(* IEC 61131-3 sources: Simulierte-Foerderanlagensteuerung/plc/function_blocks, 6 files *)

(* ---- FB_Alarm.st ---- *)
(* ============================================================================
   FB_Alarm.st
   Störmeldespeicher, Priorisierung und First-out-Erkennung.

   - Ueberlast und Not-Halt sind "lebende" Bedingungen (fallen mit dem Signal).
   - Timeout-/Stau-/Sensorstoerungen werden gespeichert und nur quittiert,
     wenn die Ursache nicht mehr ansteht.
   - eFirst haelt die zuerst aufgetretene Stoerung fest.
   ============================================================================ *)

FUNCTION_BLOCK FB_Alarm
VAR_INPUT
    xOverload            : BOOL;
    xEmergency           : BOOL;
    xStartTimeout        : BOOL;
    xStopTimeout         : BOOL;
    xJam                 : BOOL;
    xSensorInconsistency : BOOL;
    xReset               : BOOL;
END_VAR
VAR_OUTPUT
    eActive    : E_FaultCode;
    eFirst     : E_FaultCode;
    xAnyFault  : BOOL;
    xLampRed   : BOOL;
    xLampYellow: BOOL;
    xBuzzer    : BOOL;
    xOverloadLatched  : BOOL;
    xEmergencyLatched : BOOL;
    xStartLatched     : BOOL;
    xStopLatched      : BOOL;
    xJamLatched       : BOOL;
    xSensorLatched    : BOOL;
END_VAR

    (* --- Ereignisstoerungen speichern --- *)
    IF xOverload THEN
        xOverloadLatched := TRUE;
    END_IF;
    IF xEmergency THEN
        xEmergencyLatched := TRUE;
    END_IF;
    IF xStartTimeout THEN
        xStartLatched := TRUE;
    END_IF;
    IF xStopTimeout THEN
        xStopLatched := TRUE;
    END_IF;
    IF xJam THEN
        xJamLatched := TRUE;
    END_IF;
    IF xSensorInconsistency THEN
        xSensorLatched := TRUE;
    END_IF;

    (* --- Sammelstoerung --- *)
    xAnyFault := xOverloadLatched
                 OR xEmergencyLatched
                 OR xStartLatched
                 OR xStopLatched
                 OR xJamLatched
                 OR xSensorLatched;

    (* --- Quittung nur, wenn keine Ursache mehr ansteht --- *)
    IF xReset
       AND NOT xOverload
       AND NOT xEmergency
       AND NOT xStartTimeout
       AND NOT xStopTimeout
       AND NOT xJam
       AND NOT xSensorInconsistency THEN
        xOverloadLatched := FALSE;
        xEmergencyLatched := FALSE;
        xStartLatched := FALSE;
        xStopLatched := FALSE;
        xJamLatched := FALSE;
        xSensorLatched := FALSE;
    END_IF;

    (* --- Priorisierte Anzeige der aktiven Stoerung --- *)
    IF xEmergencyLatched THEN
        eActive := E_FaultCode.FAULT_EMERGENCY;
    ELSIF xOverloadLatched THEN
        eActive := E_FaultCode.FAULT_OVERLOAD;
    ELSIF xStartLatched THEN
        eActive := E_FaultCode.FAULT_START_TIMEOUT;
    ELSIF xStopLatched THEN
        eActive := E_FaultCode.FAULT_STOP_TIMEOUT;
    ELSIF xJamLatched THEN
        eActive := E_FaultCode.FAULT_JAM;
    ELSIF xSensorLatched THEN
        eActive := E_FaultCode.FAULT_SENSOR_INCONSISTENCY;
    ELSE
        eActive := E_FaultCode.FAULT_NONE;
    END_IF;

    (* --- First-out --- *)
    IF (eFirst = E_FaultCode.FAULT_NONE) AND xAnyFault THEN
        eFirst := eActive;
    END_IF;
    IF xReset AND NOT xAnyFault THEN
        eFirst := E_FaultCode.FAULT_NONE;
    END_IF;

    (* --- Meldeorgane --- *)
    xLampRed := xAnyFault;
    xBuzzer := xAnyFault;
    xLampYellow := (eActive = E_FaultCode.FAULT_JAM)
                   OR (eActive = E_FaultCode.FAULT_SENSOR_INCONSISTENCY);
END_FUNCTION_BLOCK

(* ---- FB_ConveyorProcess.st ---- *)
(* ============================================================================
   FB_ConveyorProcess.st
   Prozessablauf Automatikbetrieb.

   Zwei Varianten, gesteuert durch die Konstante AUTO_CONTINUOUS:
     - Bedarfsbetrieb (FALSE): Start bei Werkstueck am Einlauf, Nachlauf nach
       dem Auslauf, dann Rueckkehr nach IDLE.
     - Dauerlauf (TRUE): Start beim Aktivieren der Automatik, kein Stopp.

   Ausgaenge sind Impulse (ein Zyklus) fuer die Motorsteuerung.
   ============================================================================ *)

FUNCTION_BLOCK FB_ConveyorProcess
VAR_INPUT
    xEnable      : BOOL;   (* Automatik aktiv, READY, keine Stoerung *)
    xEntrySensor : BOOL;   (* B1 *)
    xExitSensor  : BOOL;   (* B2 *)
END_VAR
VAR_OUTPUT
    xStartPulse : BOOL;    (* Startimpuls an Motorsteuerung *)
    xStopPulse  : BOOL;    (* Stopimpuls an Motorsteuerung *)
    eState      : E_ProcessState;
END_VAR
VAR
    xEnablePrev : BOOL;
    tonRunOn    : TON;
    xRunOnCond  : BOOL;
END_VAR

    xStartPulse := FALSE;
    xStopPulse  := FALSE;

    (* Nachlauf-Timer jede Scan aufrufen; ausserhalb P_RUN_ON zuruecksetzen *)
    xRunOnCond := (eState = E_ProcessState.P_RUN_ON) AND NOT xExitSensor;
    tonRunOn(IN := xRunOnCond, PT := T_RUN_ON);

    IF NOT xEnable THEN
        IF xEnablePrev THEN
            xStopPulse := TRUE;   (* Automatik verlassen -> Band stoppen *)
        END_IF;
        eState := E_ProcessState.P_IDLE;
        xEnablePrev := FALSE;
    ELSE
        CASE eState OF
            E_ProcessState.P_IDLE :
                IF AUTO_CONTINUOUS THEN
                    IF NOT xEnablePrev THEN
                        xStartPulse := TRUE;
                    END_IF;
                    eState := E_ProcessState.P_TRANSPORT;
                ELSE
                    IF xEntrySensor THEN
                        xStartPulse := TRUE;
                        eState := E_ProcessState.P_TRANSPORT;
                    END_IF;
                END_IF;

            E_ProcessState.P_TRANSPORT :
                IF (NOT AUTO_CONTINUOUS) AND xExitSensor THEN
                    eState := E_ProcessState.P_RUN_ON;
                END_IF;

            E_ProcessState.P_RUN_ON :
                IF tonRunOn.Q THEN
                    xStopPulse := TRUE;
                    eState := E_ProcessState.P_IDLE;
                END_IF;

            ELSE
                eState := E_ProcessState.P_IDLE;
        END_CASE;
        xEnablePrev := TRUE;
    END_IF;
END_FUNCTION_BLOCK

(* ---- FB_Counter.st ---- *)
(* ============================================================================
   FB_Counter.st
   Werkstueckzaehlung.

   Gezaehlt wird am Auslauf ueber die steigende Flanke des Sensors B2.
   Begruendung: Der Auslauf repraesentiert ein fertig transportiertes Werkstueck.
   Die Flankenauswertung (R_TRIG) verhindert Mehrfachzaehlung, solange der
   Sensor aktiv bleibt.
   ============================================================================ *)

FUNCTION_BLOCK FB_Counter
VAR_INPUT
    xExitSensor : BOOL;    (* B2 *)
    xResetCount : BOOL;
END_VAR
VAR_OUTPUT
    diCount      : DINT;
    xJustCounted : BOOL;   (* Impuls fuer HMI/Statistik *)
END_VAR
VAR
    rtrigExit : R_TRIG;
END_VAR

    rtrigExit(CLK := xExitSensor);
    xJustCounted := FALSE;

    IF rtrigExit.Q THEN
        diCount := diCount + 1;
        xJustCounted := TRUE;
    END_IF;

    IF xResetCount THEN
        diCount := 0;
    END_IF;
END_FUNCTION_BLOCK

(* ---- FB_JamDetection.st ---- *)
(* ============================================================================
   FB_JamDetection.st
   Stau-/Blockadeerkennung.

   Verfahren: Ein Werkstueck wird am Einlauf erkannt und der Antrieb laeuft.
   Erreicht es den Auslauf nicht innerhalb T_MAX_TRANSPORT, liegt ein Stau vor.
   Die Stau-Stoerung wird bis zur Quittung gespeichert.
   ============================================================================ *)

FUNCTION_BLOCK FB_JamDetection
VAR_INPUT
    xEntrySensor      : BOOL;   (* B1 *)
    xExitSensor       : BOOL;   (* B2 *)
    xConveyorRun      : BOOL;   (* Antrieb angesteuert bzw. laeuft *)
    xReset            : BOOL;
END_VAR
VAR_OUTPUT
    xJam              : BOOL;
    xTransportPending : BOOL;   (* Werkstueck unterwegs, Auslauf erwartet *)
END_VAR
VAR
    rtrigEntry : R_TRIG;
    tonJam     : TON;
END_VAR

    rtrigEntry(CLK := xEntrySensor);

    (* Transportauftrag setzen, sobald ein Werkstueck einlaeuft und der Antrieb laeuft *)
    IF rtrigEntry.Q AND xConveyorRun THEN
        xTransportPending := TRUE;
    END_IF;

    (* Auslauf erreicht -> Transportauftrag beendet *)
    IF xExitSensor THEN
        xTransportPending := FALSE;
    END_IF;

    (* Ueberwachung der Transportzeit *)
    tonJam(IN := xTransportPending, PT := T_MAX_TRANSPORT);
    IF tonJam.Q THEN
        xJam := TRUE;
    END_IF;

    (* Quittung nur bei freiem Einlauf *)
    IF xReset AND NOT xEntrySensor THEN
        xJam := FALSE;
        xTransportPending := FALSE;
        tonJam(IN := FALSE, PT := T_MAX_TRANSPORT);
    END_IF;
END_FUNCTION_BLOCK

(* ---- FB_ModeManager.st ---- *)
(* ============================================================================
   FB_ModeManager.st
   Verwaltung der Betriebsart (Hand / Automatik).

   Der Wahlschalter ist ein reines Bedienelement; er hat keine Sicherheitsfunktion.
   ============================================================================ *)

FUNCTION_BLOCK FB_ModeManager
VAR_INPUT
    xAuto : BOOL;   (* S5: 1 = Automatik, 0 = Hand *)
END_VAR
VAR_OUTPUT
    eMode       : E_Betriebsart;
    xAutoActive : BOOL;
    xHandActive : BOOL;
END_VAR

    IF xAuto THEN
        eMode := E_Betriebsart.BETRIEB_AUTO;
    ELSE
        eMode := E_Betriebsart.BETRIEB_HAND;
    END_IF;

    xAutoActive := (eMode = E_Betriebsart.BETRIEB_AUTO);
    xHandActive := NOT xAutoActive;
END_FUNCTION_BLOCK

(* ---- FB_MotorControl.st ---- *)
(* ============================================================================
   FB_MotorControl.st
   Kern der Motorsteuerung (Steuerlogik).

   Konzept:
     - Start ist flankengesteuert (Taster bzw. Automatik-Startimpuls).
     - Selbsthaltung (Latch) des Laufwunsches.
     - Kickout-Bedingungen (Stop, Not-Halt, Ueberlast, fehlende Freigabe,
       Automatik-Stopimpuls) setzen die Selbsthaltung zurueck.
     - Stop hat Vorrang vor Start.
     - Der Schuetzbefehl ist zusaetzlich hart verriegelt.
     - Ueberwachung: "laeuft nicht an" und "stoppt nicht" ueber TON.
   ============================================================================ *)

FUNCTION_BLOCK FB_MotorControl
VAR_INPUT
    xStartManual     : BOOL;   (* S1 Start-Taster (Hand) *)
    xAutoStartPulse  : BOOL;   (* Startimpuls aus dem Automatikprozess *)
    xAutoStopPulse   : BOOL;   (* Stopimpuls (Nachlauf beendet) *)
    xStop            : BOOL;   (* TRUE = Stop betaetigt bzw. Betriebsartwechsel *)
    xEmergencyActive : BOOL;   (* Not-Halt aktiv *)
    xOverloadActive  : BOOL;   (* Ueberlast aktiv *)
    xPermissive      : BOOL;   (* Sammelfreigabe (keine Stoerung) *)
    xMotorFeedback   : BOOL;   (* tatsaechlicher Motorlauf *)
END_VAR
VAR_OUTPUT
    xContactorCmd      : BOOL; (* Befehl an Schuetz K1 *)
    xRunRequest        : BOOL; (* interne Selbsthaltung *)
    xRunning           : BOOL; (* Motor laeuft (Rueckmeldung) *)
    xFaultStartTimeout : BOOL; (* "laeuft nicht an" *)
    xFaultStopTimeout  : BOOL; (* "stoppt nicht" *)
END_VAR
VAR
    rtrigStart  : R_TRIG;
    tonStart    : TON;
    tonStop     : TON;
    xStartAction : BOOL;
    xKickout     : BOOL;
END_VAR

    (* --- Startflanke aus dem Handbetrieb --- *)
    rtrigStart(CLK := xStartManual);

    (* --- Start-/Kickout-Bedingungen --- *)
    xStartAction := (rtrigStart.Q OR xAutoStartPulse)
                    AND xPermissive
                    AND NOT xStop
                    AND NOT xEmergencyActive
                    AND NOT xOverloadActive;

    xKickout := xStop
                OR xAutoStopPulse
                OR xEmergencyActive
                OR xOverloadActive
                OR NOT xPermissive;

    (* --- Selbsthaltung des Laufwunsches; Kickout hat Vorrang --- *)
    IF xKickout THEN
        xRunRequest := FALSE;
    ELSIF xStartAction THEN
        xRunRequest := TRUE;
    END_IF;

    (* --- Schuetzbefehl, zusaetzlich hart verriegelt --- *)
    xContactorCmd := xRunRequest
                     AND NOT xStop
                     AND NOT xEmergencyActive
                     AND NOT xOverloadActive
                     AND xPermissive;

    (* --- Rueckmeldung des tatsaechlichen Motorlaufs --- *)
    xRunning := xMotorFeedback;

    (* --- Startueberwachung: Befehl EIN, keine Rueckmeldung --- *)
    tonStart(IN := xContactorCmd AND NOT xMotorFeedback,
             PT := T_MOTOR_START_TIMEOUT);
    xFaultStartTimeout := tonStart.Q;

    (* --- Stopueberwachung: Befehl AUS, Rueckmeldung bleibt EIN --- *)
    tonStop(IN := (NOT xContactorCmd) AND xMotorFeedback,
            PT := T_MOTOR_STOP_TIMEOUT);
    xFaultStopTimeout := tonStop.Q;
END_FUNCTION_BLOCK
